TYPE ST_Mode :
STRUCT
	iActMode: E_WorkingMode;
	bSetManual: BOOL;
	bSetSemi: BOOL;
	bSetAuto: BOOL;

	eModeZone:E_ModeZone:=E_ModeZone.eNone;
	
	bStateSafe_mode: BOOL:=TRUE;

END_STRUCT
END_TYPE

(* stored: Version 1.1.0.1, ProductVersion 3.1.4024.13
   DUT ST_Mode: Id {5ffe0d9a-df45-4cfe-b52b-5039f0e8974b} *)
